DATA_BLOCK "GDB_GRAPH_RecoveryTest"
{ S7_Optimized_Access := 'TRUE' }
VERSION : 0.1
NON_RETAIN
"FB_GRAPH_RecoveryTest"
BEGIN
END_DATA_BLOCK
